(* IEC 61131-3 sources: Caravan/Archiv/12-04-19/Stations/MachineControl/MachineControl/Class/Level_Class, 1 file *)

(* ---- Level_Class.st ---- *)
(*!
<Class
	Name               = "Level_Class"
	Revision           = "0.0"
	RealtimeTask       = "false"
	CyclicTask         = "true"
	DefCyclictime      = "50 ms"
	BackgroundTask     = "false"
	Sigmatek           = "false"
	OSInterface        = "false"
	HighPriority       = "false"
	Automatic          = "false"
	UpdateMode         = "Prescan"
	SharedCommandTable = "true"
	Objectsize         = "(570,240)">
	<Channels>
		<Server Name="ClassSvr" Visualized="false" Initialize="false" WriteProtected="true" Retentive="false"/>
		<Server Name="Level_X_S" Visualized="true" Remotely="true" Initialize="false" WriteProtected="false" Retentive="false"/>
		<Server Name="Level_Y_S" Visualized="true" Remotely="true" Initialize="false" WriteProtected="false" Retentive="false"/>
		<Server Name="SetZero_S" Visualized="true" Remotely="true" Initialize="false" WriteProtected="false" Retentive="false"/>
		<Server Name="ZeroPositionX_S" Visualized="true" Remotely="true" Initialize="false" WriteProtected="false" Retentive="File"/>
		<Server Name="ZeroPositionY_S" Visualized="true" Remotely="true" Initialize="false" WriteProtected="false" Retentive="File"/>
		<Client Name="PositionInput_X_C" Required="true" Internal="false"/>
		<Client Name="PositionInput_Y_C" Required="true" Internal="false"/>
	</Channels>
</Class>
*)
Level_Class : CLASS
  //Servers:
	ClassSvr 	: SvrChCmd_DINT;
	Level_X_S 	: SvrCh_DINT;
	Level_Y_S 	: SvrCh_DINT;
	ZeroPositionX_S 	: SvrCh_DINT;
	ZeroPositionY_S 	: SvrCh_DINT;
	SetZero_S 	: SvrCh_DINT;
  //Clients:
	PositionInput_X_C 	: CltCh_DINT;
	PositionInput_Y_C 	: CltCh_DINT;
  //Variables:
  //Functions:

	FUNCTION VIRTUAL GLOBAL CyWork
		VAR_INPUT
			EAX 	: UDINT;
		END_VAR
		VAR_OUTPUT
			state (EAX) 	: UDINT;
		END_VAR;
  //Tables:
	FUNCTION @STD
		VAR_OUTPUT
			ret_code	: CONFSTATES;
		END_VAR;
	FUNCTION GLOBAL TAB @CT_;
END_CLASS;

FUNCTION VIRTUAL GLOBAL Level_Class::CyWork
	VAR_INPUT
		EAX 	: UDINT;
	END_VAR
	VAR_OUTPUT
		state (EAX) 	: UDINT;
	END_VAR

    //Einlesen
    PositionInput_X_C   :=      PositionInput_X_C.Read();
    PositionInput_Y_C   :=      PositionInput_Y_C.Read();

    //Nullpunkt definieren
    if SetZero_S  = 1 then

      ZeroPositionX_S :=  ZeroPositionX_S.Write(input:=PositionInput_X_C);
      ZeroPositionY_S :=  ZeroPositionY_S.Write(input:=PositionInput_Y_C);

    end_if;

    //Lage für X Achse ausgeben
    Level_X_S   :=    (PositionInput_X_C - ZeroPositionX_S + 310) ;

    //Nicht übersteuern, im Bildausschnitt bleiben
    IF Level_X_S  > 619  THEN

       Level_X_S   :=    Level_X_S.Write(input:=619);

    ELSIF    Level_X_S  < 1 THEN

        Level_X_S   :=    Level_X_S.Write(input:=1);

    ELSE

        Level_X_S   :=    Level_X_S.Write(input:=Level_X_S);

    END_IF;

    //Lage für die Y Achse ausgeben
    Level_Y_S   :=    PositionInput_Y_C - ZeroPositionY_S +165;

    //Nicht übersteuern, im Bildausschnitt bleiben
    IF Level_Y_S > 329 THEN

      Level_Y_S   :=  Level_Y_S.Write(input:=329);

    ELSIF   Level_Y_S < 1 Then

             Level_Y_S  :=  Level_Y_S.Write(input:=1);

    ELSE

      Level_Y_S   :=    Level_Y_S.Write(input:=Level_Y_S);

    END_IF;

	state := READY;

END_FUNCTION
